{attribute 'qualified_only'}
{attribute 'strict'}
{attribute 'to_string'}
TYPE XtsResetState :
(
	Idle := 0,
	ResettingHardware := 1,
	ResettingCAGroup := 2,
	Done
);
END_TYPE

(* stored: Version 1.1.0.1
   DUT XtsResetState: Id {dd747b37-d26a-4058-8f31-1a51dab41710} *)
